Staubli VAL3: sPointTemplate.dtx

public bool bActive
public pointRx pPointRx = {fatherId=world[0]}
public string sName
